Fanuc KAREL source: KT00683.KL

PROGRAM KT00683
%NOLOCKGROUP
VAR
  P1: JOINTPOS
  P2: JOINTPOS
  OUT: REAL
BEGIN
  OUT = + P1
END KT00683
